(* IEC 61131-3 sources: TSA-FMICS22/ahorn/test/lib_pass/file/ssa, 2 files *)

(* ---- parts_of_antivalent.st ---- *)
PROGRAM P
VAR_INPUT
    Activate       : BOOL := FALSE;
END_VAR
VAR
    Ready          : BOOL := FALSE;
    S_TwoHandOut   : BOOL := FALSE;
    DiagCode       : WORD := 16#0;
END_VAR
    IF NOT Activate THEN
        DiagCode := 16#0000;
    ELSE
     CASE DiagCode OF
     16#0000:
         IF Activate THEN
              DiagCode := 16#8001;
         END_IF;
     END_CASE;
    END_IF;

    CASE DiagCode OF
    16#0000:
        Ready := FALSE;
        S_TwoHandOut := FALSE;
    16#8000:
        Ready := TRUE;
        S_TwoHandOut := TRUE;
    16#8001:
        Ready := TRUE;
        S_TwoHandOut := FALSE;
    END_CASE;
END_PROGRAM

(* ---- wikipedia_example.st ---- *)
PROGRAM P
VAR
    w : INT;
    x : INT;
    y : INT;
    z : INT;
END_VAR
    x := 5;
    x := x - 3;
    IF x < 3 THEN
        y := x * 2;
        w := y;
    ELSE
        y := x - 3;
    END_IF;
    w := x - y;
    z := x + y;
END_PROGRAM
